Staubli VAL3: ParaItem.dtx

public mdesc mMdesc
public num nMoveType
public num nActionIndex
public num nPercentage
public ifItem iIfItem
  [0]
    num nSigType[3]
    num nSigIndex[3]
    num nValue[3]
    bool bANDOR[2]
public num nDelay
public num nSigValue
public bool bSafePoint
